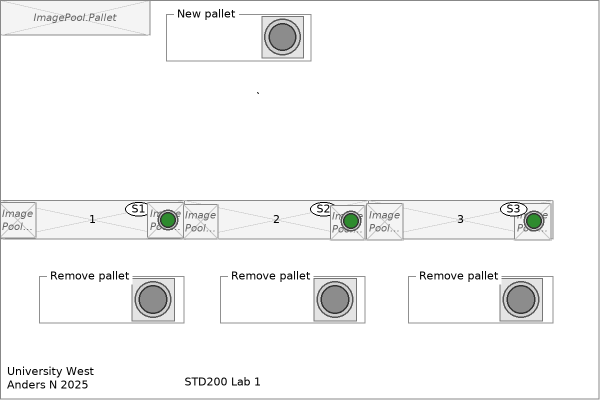
VISUALIZATION Visualization  // 600x400
    Label (4,363 125x30), "University West Anders N 2025"
    Image (0,200 185x39), "1", image: ImagePool.Conveyor
    Image (184,200 185x39), "2", image: ImagePool.Conveyor
    Image (368,200 185x39), "3", image: ImagePool.Conveyor
    Image (0,0 150x35), image: ImagePool.Pallet
        p3560616238: MAIN.miPallet1PosX
        p2738717112: MAIN.miPallet1PosY
    Image (0,0 150x35), image: ImagePool.Pallet
        p3560616238: MAIN.miPallet2PosX
        p2738717112: MAIN.miPallet2PosY
    Image (0,0 150x35), image: ImagePool.Pallet
        p3560616238: MAIN.miPallet3PosX
        p2738717112: MAIN.miPallet3PosY
    Image (514,203 37x37), invisible if: NOT MAIN.mxMotor3Running, image: ImagePool.Rotate
    Ellipse (125,202 27x14), "S1", tooltip "Sensor 1", colour toggle: MAIN.qxSensor1
    Ellipse (310,202 27x14), "S2", tooltip "Sensor 2", colour toggle: MAIN.qxSensor2
    Ellipse (500,202 27x14), "S3", tooltip "Sensor 3", colour toggle: MAIN.qxSensor3
    PushSwitch (497,278 48x43), tooltip "Empty Conveyor 3", variable: MAIN.mxEmptyConvayor3, behaviour: TAP, style: Switch-PushSwitch-Gray
    PushSwitch (311,278 48x43), tooltip "Empty Conveyor 2", variable: MAIN.mxEmptyConvayor2, behaviour: TAP, style: Switch-PushSwitch-Gray
    PushSwitch (129,278 48x43), tooltip "Empty Conveyor 1", variable: MAIN.mxEmptyConvayor1, behaviour: TAP, style: Switch-PushSwitch-Gray
    Image (-1,202 37x36), invisible if: NOT MAIN.mxMotor1Running, image: ImagePool.Rotate
    Image (147,202 37x36), invisible if: NOT MAIN.mxMotor1Running, image: ImagePool.Rotate
    Image (183,204 35x35), invisible if: NOT MAIN.mxMotor2Running, image: ImagePool.Rotate
    Image (330,205 35x35), invisible if: NOT MAIN.mxMotor2Running, image: ImagePool.Rotate
    Image (366,203 37x37), invisible if: NOT MAIN.mxMotor3Running, image: ImagePool.Rotate
    Label (99,363 251x38), "STD200 Lab 1"
    Polyline (257,92) (258,93)
    Lamp1 (155,208 26x24), variable: MAIN.mxMotor1Running, style: Lamp-Lamp1-Green
    Lamp1 (338,209 26x24), variable: MAIN.mxMotor2Running, style: Lamp-Lamp1-Green
    Lamp1 (521,209 26x24), variable: MAIN.mxMotor3Running, style: Lamp-Lamp1-Green
    Label (198,6 87x21)
    GroupBox (39,268 145x55), "Remove pallet"
    GroupBox (220,268 145x55), "Remove pallet"
    GroupBox (408,268 145x55), "Remove pallet"
    GroupBox (166,6 145x55), "New pallet"
        PushSwitch (94,10 45x42), tooltip "Load a pallet", variable: MAIN.mxLoadPallet, behaviour: TAP, style: Switch-PushSwitch-Gray
END_VISUALIZATION

(* stored: Version 1.1.0.1
   Visu Visualization: Id {ad45f26b-89f6-408d-b081-64ca21bca6cc} *)
